Yaskawa INFORM job: 0523.JBI

/JOB
//NAME 0523
///FOLDERNAME FOLDER004
//POS
///NPOS 18,0,0,0,0,0
///TOOL 1
///POSTYPE PULSE
///PULSE
C00000=-1,-38943,-47654,0,-74515,0
C00001=-41491,4068,-52360,6325,-57867,-68771
C00002=-42127,24040,-59211,-18,-27953,-66868
C00003=-42899,24480,-58538,-44,-28085,-66613
C00004=-48638,32602,-45619,-1836,-31314,-44796
C00005=-47067,42694,-28404,-2184,-36429,-26338
C00006=-45244,46402,-21808,-2097,-38148,-26966
C00007=-39546,54387,-7194,-1554,-43041,-9553
C00008=-32482,55159,-5756,-685,-43914,5330
C00009=-27698,52425,-10834,-806,-42445,3862
C00010=-18800,45607,-23229,826,-39050,25331
C00011=-16780,36282,-39470,2017,-34318,42079
C00012=-17583,32074,-46479,2118,-32649,42278
C00013=-26276,20156,-65020,2085,-27338,74127
C00014=-34910,20741,-64159,400,-27049,92913
C00015=-35627,21061,-63687,375,-27132,93151
C00016=-40407,-9140,-58390,121,-53542,94785
C00017=-1,-38943,-47654,0,-74515,0
//INST
///DATE 2018/05/22 20:35
///ATTR SC,RW
///GROUP1 RB1
NOP
MOVJ C00000 VJ=30.00
MOVJ C00001 VJ=30.00
MOVL C00002 V=133.3
MOVL C00003 V=10.0
MOVL C00004 V=10.0
MOVL C00005 V=10.0
MOVL C00006 V=10.0
MOVL C00007 V=10.0
MOVL C00008 V=10.0
MOVL C00009 V=10.0
MOVL C00010 V=10.0
MOVL C00011 V=10.0
MOVL C00012 V=10.0
MOVL C00013 V=10.0
MOVL C00014 V=10.0
MOVL C00015 V=10.0
MOVL C00016 V=133.3
MOVJ C00017 VJ=30.00
END
